// TwinCAT 3 PLC project PLCStudent
// ProgramVersion: 3.1.4026.20
// libraries:
//   Tc2_Standard, * (Beckhoff Automation GmbH)
//   Tc2_System, * (Beckhoff Automation GmbH)
//   Tc3_Module, * (Beckhoff Automation GmbH)
// project tree:
//   GVLs/ GVL.TcGVL
//   / PlcTask.TcTTO
//   POUs/ MAIN.TcPOU, Control_FBD.TcPOU
// (motion and I/O tree: see PLC project plcsim)
// real-time tasks:
//   TASK PlcTask: cycle T#80ms, priority 1, ADS port 350
//   TASK PlcTask1: cycle T#10ms, priority 20, ADS port 351
// variable links:
//   PLCSim/PLCSim Instance <-> PLCStudent/PLCStudent Instance
//     PlcTask Inputs/MAIN.ixRunConveyor1 <-> PlcTask Outputs/Control_FBD.qxRunConveyor1
//     PlcTask Inputs/MAIN.ixRunConveyor2 <-> PlcTask Outputs/Control_FBD.qxRunConveyor2
//     PlcTask Inputs/MAIN.ixRunConveyor3 <-> PlcTask Outputs/Control_FBD.qxRunConveyor3
//     PlcTask Outputs/MAIN.qxSensor1 <-> PlcTask Inputs/Control_FBD.ixSensor1
//     PlcTask Outputs/MAIN.qxSensor2 <-> PlcTask Inputs/Control_FBD.ixSensor2
//     PlcTask Outputs/MAIN.qxSensor3 <-> PlcTask Inputs/Control_FBD.ixSensor3

CONFIGURATION PLCStudent
    RESOURCE PLC ON TwinCAT3
        TASK PlcTask(INTERVAL := T#10ms, PRIORITY := 20);
        PROGRAM MAIN WITH PlcTask : MAIN;
    END_RESOURCE
END_CONFIGURATION

// ---- GVLs/GVL.TcGVL
{attribute 'qualified_only'}
VAR_GLOBAL	


END_VAR

// ---- POUs/MAIN.TcPOU
PROGRAM MAIN
VAR
END_VAR

Control_FBD();

END_PROGRAM

// ---- POUs/Control_FBD.TcPOU
PROGRAM Control_FBD
VAR
	ixSensor1		AT %I*:	BOOL; 		//Pallet on sensor1 (S1)
	ixSensor2		AT %I*:	BOOL; 		//Pallet on sensor2 (S2)
	ixSensor3		AT %I*:	BOOL; 		//Pallet on sensor3 (S3)

	qxRunConveyor1	AT %Q*:	BOOL; 		// Motor that runs Conveyor 1*)
	qxRunConveyor2	AT %Q*:	BOOL; 		// Motor that runs Conveyor 2*)
	qxRunConveyor3	AT %Q*:	BOOL; 		// Motor that runs Conveyor 3*)	

	//Transport memory
	mxTrpConveyor1to2 : BOOL;
	mxTrpConveyor2to3 : BOOL;

END_VAR

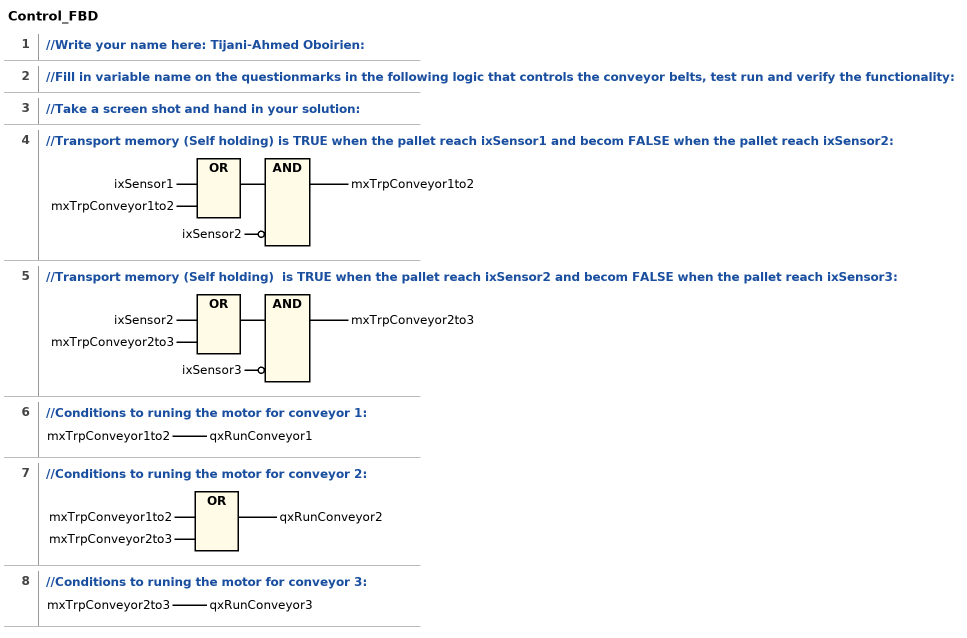
// NETWORK 1
// label: //Write your name here: Tijani-Ahmed Oboirien

// NETWORK 2
// label: //Fill in variable name on the questionmarks in the following logic that controls the conveyor belts, test run and verify the functionality

// NETWORK 3
// label: //Take a screen shot and hand in your solution

// NETWORK 4
// label: //Transport memory (Self holding) is TRUE when the pallet reach ixSensor1 and becom FALSE when the pallet reach ixSensor2
mxTrpConveyor1to2 := (ixSensor1 OR mxTrpConveyor1to2) AND NOT ixSensor2;

// NETWORK 5
// label: //Transport memory (Self holding)  is TRUE when the pallet reach ixSensor2 and becom FALSE when the pallet reach ixSensor3
mxTrpConveyor2to3 := (ixSensor2 OR mxTrpConveyor2to3) AND NOT ixSensor3;

// NETWORK 6
// label: //Conditions to runing the motor for conveyor 1
qxRunConveyor1 := mxTrpConveyor1to2;

// NETWORK 7
// label: //Conditions to runing the motor for conveyor 2
qxRunConveyor2 := mxTrpConveyor1to2 OR mxTrpConveyor2to3;

// NETWORK 8
// label: //Conditions to runing the motor for conveyor 3
qxRunConveyor3 := mxTrpConveyor2to3;

END_PROGRAM
